Fanuc KAREL source: kt00490.KL

PROGRAM KT00490
%STACKSIZE=65535
%PRIORITY=65535
%NOLOCKGROUP
VAR
P1 : POSITION
P2 : JOINTPOS9
OUT : XYZWPR
BEGIN
-- UNRESOLVED_PC line 8 opcodes [49 49 7E 60 7E 4A] marker_code=0
END KT00490
